ABB RAPID module: TgtProg.mod

MODULE MainModule

GLOBAL Proc main()
    TPWrite "m "q" ";
    ab(cd);
    xy;
    raw code
EndProc
EndModule
